// TIA Portal V20 export
// export: Created 2026-10-20T18:55:40.6540563Z, ExportSetting None, DisplayName Totally Integrated Automation Portal, DisplayVersion V20 Update 6, DisplayName TIA Portal Openness, DisplayVersion V20 Update 6, DisplayName TIA Portal Version Control Interface, DisplayVersion V20 Update 6, DisplayName SINAMICS Startdrive Advanced, DisplayVersion V20 SP1, DisplayName SINAMICS Startdrive G130, G150, S120, S150, SINAMICS MV, G220, S200, S210, DisplayVersion V20 SP1, DisplayName SINAMICS Startdrive G110M, G120, G120C, G120D, G120P, G115D, DisplayVersion V20 SP1, DisplayName STEP 7 Professional, DisplayVersion V20 Update 6, DisplayName STEP 7 Safety, DisplayVersion V20 Update 2, DisplayName WinCC Basic/Comfort/Advanced, DisplayVersion V20 Update 6, DisplayName WinCC Unified, DisplayVersion V20 Update 6
VAR_GLOBAL   // PLC tag table "Lock_1"
   Lock_1_Estop_CH2 AT %I1758.3 : Bool;
   Lock_1_Closed_CH2 AT %I1758.1 : Bool;
   Lock_1_Closed_CH1 AT %I1758.0 : Bool;
   Lock_1_Estop_CH1 AT %I1758.2 : Bool;
   "Solenoid Enable_1" AT %Q766.0 : Bool;
   Lamps_1 AT %QB369 : Byte;
   Lock_1_Reset_Input2 AT %Q1759.1 : Bool;
   Lock_1_Reset_Input4 AT %Q1759.3 : Bool;
   Lock_1_Reset_Input3 AT %Q1759.2 : Bool;
   Switches_1 AT %IB142 : Byte;
   Lock_1_Reset_Input1 AT %Q1759.0 : Bool;
   "Lock Reset_1" AT %Q767.0 : Bool;
   "Lock Position_1" AT %I204.0 : Bool;
   "Guard Position_1" AT %I143.0 : Bool;
END_VAR
